(* IEC 61131-3 sources: vscode-twincat-st/src/sample, 1 file *)

(* ---- stubs.st ---- *)
// ADR delivers the address of its argument in a PVOID
FUNCTION ADR : PVOID

END_FUNCTION
